(* IEC 61131-3 sources: daoli-st-library/DL_Process (part 67) *)

(* ---- FB_DL_ModbusPollMaster.st ---- *)
(*==============================================================================
 * 组件名称 (Component)  : FB_DL_ModbusPollMaster
 * 所属子库 (Sublibrary) : DL_Process
 * 当前版本 (Version)    : 1.0.0
 * 分类     (Category)   : 通信调度功能块（Function Block · 轮询主站调度抽象层）
 * 作者     (Author)     : Daoli Library
 * 日期     (Date)       : 2026-11-15
 * 兼容性   (Platform)   : CODESYS 3.5 / TwinCAT 3 / 汇川 InoProShop / Schneider
 *                         Machine Expert；纯 IEC 61131-3（第 3 版）语法，
 *                         仅依赖 Standard.library（TON / F_TRIG），零厂商方言
 * 功能简介 (Function)   : 多从站轮询主站调度器（Modbus RTU 轮询节拍抽象层）。
 *                         按站表顺序轮询、单事务响应超时重试、成功/异常双计数器
 *                         台账、空表与全跳过保护、站表禁用跳过的自动回绕。本块
 *                         只做「调度」：决定「此刻该问哪个站、问什么地址区、失败
 *                         重试几次、超时怎么记账」，帧的构造、CRC 校验、字节收发、
 *                         串口/TCP 底层时序全部交由传输层实现。
 * 分层声明 (Layering)   : ① 本块不绑定任何具体串口库、不引用任何厂商驱动块；
 *                         ② 传输层经两个抽象方法 SendFrame / RecvFrame 由集成者
 *                         实现（推荐做法：EXTENDS 本块并覆盖 DoTransaction 作为
 *                         统一入口，在覆盖体内调用自家收发库，再复用本块的记账
 *                         与重试；亦可只覆盖 SendFrame / RecvFrame 两个帧级原语）；
 *                         ③ 基类默认实现为「抽象桩」：返回 FALSE 并锁故障码
 *                         0005_0290（传输层未实现），这是抽象层的合法形态，不是
 *                         漏填——未注入传输层时块不会静默假成功；
 *                         ④ 调度层零触碰帧内容：不解析功能码、不读写应答字节、
 *                         不做 CRC 运算。CRC-16/Modbus 的公开算法定义在本库已有
 *                         实现（见 DL_MathData 子库既有 CRC 计算函数），本块仅在
 *                         此注释说明「可作校验实现」，不 import、不调用、不内联。
 * 职责边界 (Scope)      : ① 不做站内数据解包与工程量换算（由上层按站表项自行
 *                         读取应答缓冲后处理）；② 不做主备链路切换与总线诊断
 *                         （后续轮次另立组件）；③ 不做写单寄存器/写多寄存器的
 *                         流程编排（功能码仅作透传字段，调度节拍与读写无关）。
 * 开源溯源 (Origin)     : 来源标签 codesys-forge-modbus（T1-4 开族续挖）。仅参考
 *                         CODESYS Forge 免费库 ModbusFB 公开文档页中「主站轮询 /
 *                         站表组织 / 超时重试 / 轮询间隔」的功能分类与参数域惯例，
 *                         以及「帧构造与校验归传输层」的分层语义；所据页面未显
 *                         式声明许可条款，故按最严口径处置：只借组织分类与参数
 *                         范围，零代码行复制。本块的枚举编号、状态机、站表结构、
 *                         台账口径与故障码位 100% 本库独立设计，clean-room 实现。
 * 公约遵循 (Convention) : 0.1/R19 首扫范式（IF (NOT _bInit)）；0.2/R21 bError 显式
 *                         排除信息级码；0.5/R7 定时器与边沿实例主体最前部无条件
 *                         刷新；0.6/R14 定时器语义参数变化断输入一拍；0.7/R15 故障
 *                         级锁存仅重建路径清码；0.9 出口默认值先赋；0.14 WHILE 带
 *                         防死锁计数器 + 数组访问先判上下界；0.16 阈值全常量化。
 * 红线自检 (Redline)    : 全局隔离 ✓（零全局变量表引用、零外部变量声明、零物理
 *                         地址字面记号）｜命名合规 ✓（b/n/u/f/t/a/st/e/fb/i 前缀
 *                         全覆盖）｜注释完整 ✓（声明行 100% 中英双语同行注释）｜
 *                         OOP 封装 ✓（内部状态全私有，传输层经抽象方法注入）｜
 *                         周期安全 ✓（TON / F_TRIG 实例无条件刷新，方法无跨周期
 *                         驻留）｜防御编程 ✓（索引判界、循环防死锁、重试上限、
 *                         ENUM + CASE + ELSE 兜底）｜可移植性 ✓（纯 IEC 61131-3）｜
 *                         终结符成对 ✓
 * 设计要点 (Key notes)  : ① 事务生命周期：eRequest 发起（一次性调用抽象方法）→
 *                         eWaitResp 轮询结果（ePending 等待、eDone 成功、
 *                         eTimeout/eFailed 失败）→ eSttUpdate 记账 → eNextStn。
 *                         传输层可为异步（返回 FALSE 且 eResult = ePending 表示
 *                         尚未收完），调度层的响应超时定时器是它的兜底下限。
 *                         ② 不因单站失败中断轮询：重试耗尽只累加该站异常计数并
 *                         继续下一站（台账留证，避免一站坏总线导致全线停摆）；
 *                         只有「传输层未实现」与「站表索引越界」才锁全局故障。
 *                         ③ 轮询间隔由 TON 闸门实现（eSttUpdate 后重新计时），
 *                         事务结束到下一次发起至少间隔 tPollInterval，防止从站
 *                         换向静默期被打断（RTU 帧间静默的工程近似）。
 *                         ④ 站表回绕：每次事务结束把索引 +1，寻找下一站时从当前
 *                         索引起最多检查 uStationCount 站（超过即回绕），全部
 *                         跳过则置信息级码并按间隔节流空转，不锁故障。
 *                         ⑤ 计数口径：uStatOk / uStatErr 累计在调用方持有的站表
 *                         项内（跨班不清零），本块自身不保存历史，重启即从站表
 *                         现值继续，便于 HMI 做长期台账。
 * 偏离留档 (Deviation)  : ① 规格建议故障码 0005_0290~0293 中 0293 未使用（站数
 *                         非法按钳位 + 信息级处置，不锁故障；理由：站数是可在线
 *                         修改的组态量，钳位比停机更符合现场），实际使用
 *                         0005_0290~0292 三条；
 *                         ② 传输层抽象未采用独立 INTERFACE 文件（理由：本库公约
 *                         0.18「一文件一 POU」，接口件须独立成 .st 且本泳道不
 *                         允许新增第 6 个文件；改为块内抽象方法三件套，语义等价：
 *                         基类桩返回 FALSE + 锁码，派生块覆盖实现）；
 *                         ③ 规格 VAR 段 bFirstScan 改名 _bInit（公约 0.1 统一命名）。
 * 故障码表 (Error codes) :
 *                         16#0005_0190【信息级】站数越界已钳位到 1 至 16
 *                         16#0005_0191【信息级】站表全部跳过，本轮无事务（按间隔节流）
 *                         16#0005_0192【信息级】单站重试耗尽，异常台账已累加
 *                         16#0005_0193【信息级】超时/间隔参数非法已兜底
 *                         16#0005_0290【故障级】传输层未实现（抽象方法桩未被覆盖）
 *                         16#0005_0291【故障级】站表索引越界（越界保护触发）
 *                         16#0005_0292【故障级】非法状态兜底（枚举越界）
 * 验收向量 (Acceptance) :
 *   V1 单站成功：站数 1、从站 1 功能码 3 → eRequest 发起一次，eWaitResp 得
 *      eDone → uStatOk +1、bDone 单拍、回到 eNextStn；
 *   V2 超时重试：传输层持续回 ePending → 响应超时定时器到期后 uActiveRetry
 *      逐次 +1，达 uMaxRetry 后该站 uStatErr +1 且轮询继续下一站（不锁故障）；
 *   V3 站表跳过：站 0 的 bSkip = TRUE → 首个事务直接落在站 1（索引回绕正确）；
 *      全部站跳过 → 信息级 0191，块按 tPollInterval 节流空转，bBusy FALSE；
 *   V4 抽象桩：未覆盖 DoTransaction / SendFrame / RecvFrame → 首次发起即锁
 *      0005_0290 并停轮询，bError TRUE（杜绝静默假成功）；
 *   V5 间隔节流：tPollInterval = 100 ms、任务 10 ms → 相邻两事务发起间隔
 *      不少于 100 ms（TON 闸门计时）；
 *   V6 禁用重建：bEnable 下降沿 → 队伍暂停且保持现场（站索引/计数不清零），
 *      再次使能从原索引继续，不重复打扰刚问过的站。
 * 修订历史 (Revision)   :
 *   2026-11-15  v1.0.0  首版入库（Round 09 · DL_Process Modbus 轮询调度件）
 *============================================================================*)

(*-----------------------------------------------------------------------------
 * 集成示例 (Integration guide)：
 *   1 定义派生块 FB_MyRtuMaster EXTENDS FB_DL_ModbusPollMaster，覆盖
 *     DoTransaction（VAR_IN_OUT stItem : ST_DL_PollItem），在覆盖体内调用自家
 *     串口收发块完成「组帧 + 发送 + 收帧 + CRC 校验」，并把结果写回本块事务
 *     上下文（成功回 eDone，超时回 eTimeout，异常码回 uExceptionCode）。
 *   2 上层每周期调用派生块实例，注入站表数组与调度参数：
 *      aPollTable[0].uSlaveAddr := 1; aPollTable[0].uFuncCode := 3;
 *      aPollTable[0].uStartAddr := 0; aPollTable[0].uQuantity := 16;
 *      fbPoll(uStationCount := 4, tRespTimeout := T#500MS, uMaxRetry := 3,
 *             tPollInterval := T#100MS, aPollTable := aPollTable);
 *   3 读台账：aPollTable[i].uStatOk / uStatErr 由本块维护，HMI 直接读结构体。
 *----------------------------------------------------------------------------*)

(*-----------------------------------------------------------------------------
 * 常见误用与现场提示 (Field notes)：
 *   1 站表项的功能码只是透传字段，本块不校验其合法性；上位填 0 或非法功能码
 *     时，从站会回异常码，表现为该站 uStatErr 持续上升，请查站表而不是本块。
 *   2 响应超时必须大于最慢从站的最长应答时间；填得过小会造成「其实成功但被
 *     判超时」的重复点名，从站可能因此回异常码（上一次未收完）。
 *   3 uMaxRetry = 0 表示不重试，一次失败即记账进下一站，适合「宁漏不拖」的
 *     快速巡检场景。
 *   4 站表全部 bSkip 时本块按间隔空转且 bBusy 恒 FALSE，这是正常状态，不是
 *     死机；检修期整线隔离时常被误判为故障。
 *   5 本块不做总线抢占仲裁：同一物理链路上不要挂两个本块实例，否则帧会交错。
 *----------------------------------------------------------------------------*)

(*-----------------------------------------------------------------------------
 * 枚举: E_DL_PollState（归属 FB_DL_ModbusPollMaster，随本文件发布）
 * 含义: 轮询调度离散状态。数值步长 10 留空位，故障态 99 保证排序末位。
 *----------------------------------------------------------------------------*)
{attribute 'strict'}
{attribute 'qualified_only'}
TYPE E_DL_PollState :
(
    eIdle      := 0,     // 空闲：未使能或故障重建后待启动 / Idle: disabled or waiting for a rebuild
    eNextStn   := 10,    // 选下一站：按站表回绕寻找未跳过站，并受轮询间隔闸门约束 / Select next station with wrap and interval gating
    eRequest   := 20,    // 发起事务：一次性调用抽象方法 DoTransaction / Issue one transaction by calling DoTransaction
    eWaitResp  := 30,    // 等待应答：轮询传输层结果与响应超时定时器 / Wait for the transport result and the response timeout
    eSttUpdate := 40,    // 记账：成功/异常计数累加并产生单拍完成脉冲 / Accounting with a one-scan done pulse
    eFault     := 99     // 故障锁存：仅使能下降沿重建可退 / Fault latched, left only by the disable-edge rebuild
) UINT;
END_TYPE

(*-----------------------------------------------------------------------------
 * 枚举: E_DL_MbTxnResult（归属 FB_DL_ModbusPollMaster，随本文件发布）
 * 含义: 单事务结果，由传输层回填。调度层只据此推进状态，不解析帧内容。
 *----------------------------------------------------------------------------*)
{attribute 'strict'}
{attribute 'qualified_only'}
TYPE E_DL_MbTxnResult :
(
    ePending := 0,       // 传输中：尚未收完应答（异步传输层的等待态） / In progress, response not yet complete
    eDone    := 10,      // 事务成功：应答完整且通过传输层校验 / Success, a complete and validated response
    eTimeout := 20,      // 传输超时：传输层自身判超时 / Timeout reported by the transport layer
    eFailed  := 30       // 传输失败：校验错、异常码或链路错误 / Failure such as a check error, an exception or a link error
) UINT;
END_TYPE

(*-----------------------------------------------------------------------------
 * 结构体: ST_DL_PollItem（归属 FB_DL_ModbusPollMaster，随本文件发布）
 * 用途: 站表项。由调用方持有并注入（VAR_IN_OUT 数组），本块只读写统计字段。
 * 说明: uFuncCode / uStartAddr / uQuantity 均为透传字段，本块不解析、不改写。
 *----------------------------------------------------------------------------*)
TYPE ST_DL_PollItem :
STRUCT
    uSlaveAddr : USINT := 1;      // 从站地址（Slave address）[1~247]，0 与 248 以上为保留地址 / Reserved above 247 and at zero
    uFuncCode  : USINT := 3;      // 功能码（Function code），本块仅透传不解析 / Passed through, never parsed by this block
    uStartAddr : UINT := 0;       // 起始地址（Start address），寄存器区偏移，本块仅透传 / Register offset, passed through only
    uQuantity  : UINT := 1;       // 数量（Quantity），寄存器个数或线圈个数，本块仅透传 / Register or coil count, passed through only
    uStatOk    : UDINT := 0;      // 成功计数（Success counter）[次]，跨班累计由调用方清零 / Accumulated until the caller clears it
    uStatErr   : UDINT := 0;      // 异常计数（Error counter）[次]，重试耗尽即累加 / Incremented when the retries are exhausted
    bSkip      : BOOL := FALSE;   // 本站跳过（Skip this station），TRUE 时轮询回绕绕过本站 / TRUE makes the scan wrap past this station
END_STRUCT
END_TYPE

(*-----------------------------------------------------------------------------
 * 结构体: ST_DL_ModbusTxn（归属 FB_DL_ModbusPollMaster，随本文件发布）
 * 用途: 单事务上下文。调度层装填请求字段，传输层回填结果字段，双方以此交接。
 * 说明: 应答缓冲容量 256 字节为 Modbus RTU 最大帧长度（地址 + 功能码 + 数据 +
 *       CRC 的上限），调度层只保存不解读。
 *----------------------------------------------------------------------------*)
TYPE ST_DL_ModbusTxn :
STRUCT
    uSlaveAddr     : USINT := 1;                        // 从站地址（Slave address）[1~247] / Slave address in the range one to 247
    uFuncCode      : USINT := 3;                        // 功能码（Function code），透传 / Passed-through function code
    uStartAddr     : UINT := 0;                         // 起始地址（Start address），透传 / Passed-through start address
    uQuantity      : UINT := 1;                         // 数量（Quantity），透传 / Passed-through quantity
    eResult        : E_DL_MbTxnResult := E_DL_MbTxnResult.ePending; // 事务结果（Transaction result），传输层回填 / Filled in by the transport layer
    uExceptionCode : USINT := 0;                        // 异常码（Exception code）[1~255]，0 = 无异常，传输层回填 / Zero means no exception
    uRxLen         : UINT := 0;                         // 应答字节数（Response length）[字节]，传输层回填 / Response length in bytes
    auRxFrame      : ARRAY[0..255] OF BYTE;             // 应答帧原始字节（Raw response frame）[字节]，容量 256，调度层不解读 / Raw bytes, never parsed here
    bAbort         : BOOL := FALSE;                     // 中止请求（Abort request），重试或切站时由调度层置位 / Set by the scheduler on retries
END_STRUCT
END_TYPE

(*==============================================================================
 * 功能块: FB_DL_ModbusPollMaster
 * 调用约定: 每个扫描周期无条件调用一次；站表与参数全部经引脚注入。
 * 抽象层形态: DoTransaction / SendFrame / RecvFrame 三个默认实现均为抽象桩
 *             （返回 FALSE 并锁 0005_0290），由派生块覆盖后落地真实传输。
 *============================================================================*)
FUNCTION_BLOCK FB_DL_ModbusPollMaster
VAR_INPUT
    bEnable       : BOOL;               // 调度使能（Scheduler enable），FALSE 时队列暂停并保持现场 / FALSE pauses the queue and keeps the context
    uStationCount : UINT := 4;          // 轮询站数（Station count）[站]，域 1~16，越界钳位 / Clamped to the range one to sixteen
    tRespTimeout  : TIME := T#500MS;    // 单事务响应超时（Response timeout）[ms]，域 >= 1 ms / At least one millisecond
    uMaxRetry     : UINT := 3;          // 超时重试上限（Retry limit）[次]，0 = 不重试 / Zero means no retry
    tPollInterval : TIME := T#100MS;    // 相邻事务最小间隔（Minimum poll interval）[ms]，0 = 不节流 / Zero disables the interval gate
END_VAR
VAR_OUTPUT
    bBusy          : BOOL;              // 有事务执行中（Transaction in progress）/ A transaction is running
    uActiveStation : UINT;              // 当前轮询站索引（Active station index）[索引 0~15] / Active station index in the range zero to fifteen
    uActiveRetry   : UINT;              // 当前站累计重试数（Active retry count）[次]，切站清零 / Cleared when the station advances
    bDone          : BOOL;              // 单站事务完成（Station transaction done），单拍脉冲（R25）/ One-scan pulse per station completion
    bError         : BOOL;              // 故障保持型（Fault latched），显式排除信息级码 / Latched fault flag, info codes excluded
    uErrorId       : UDINT;             // 故障码（Error code），0 = 无故障，段位 16#0005_xxxx / Error code, zero means no error
END_VAR
VAR_IN_OUT
    aPollTable    : ARRAY[0..DL_MB_MAX_STN-1] OF ST_DL_PollItem; // 轮询站表（Poll table），调用方持有 / Caller-owned poll table
END_VAR
VAR
    _eState       : E_DL_PollState := E_DL_PollState.eIdle; // 主状态机状态（Main state machine state）/ Main state machine state
    _bInit        : BOOL;               // 首扫完成标志（First-scan done flag），初值 FALSE / First-scan done flag, initial FALSE
    _uStnIdx      : UINT;               // 当前站索引（Current station index）[索引]，域 0~15 / Station index in the range zero to fifteen
    _uRetryCnt    : UINT;               // 重试计数（Retry counter）[次] / Retry counter
    _uStnCntEff   : UINT := 4;          // 生效站数（Effective station count）[站]，钳位后 / Effective station count after clamping
    _uStnTried    : UINT;               // 已检查站数（Stations examined）[站]，回绕寻找用 / Stations examined during the wrap search
    _uGuard       : UINT;               // 循环防死锁计数（Loop guard counter）[次]，上限 16 / Loop guard bounded by sixteen
    _bStationFound : BOOL;              // 找到可轮询站（Usable station found）/ A usable station was found
    _tRespEff     : TIME := T#500MS;    // 生效响应超时（Effective response timeout）[ms] / Effective response timeout [ms]
    _tGapEff      : TIME := T#100MS;    // 生效轮询间隔（Effective poll interval）[ms] / Effective poll interval [ms]
    _bGapActive   : BOOL;               // 间隔闸门激活（Interval gate armed），TRUE 时须等定时器到期 / The gate holds until the timer elapses
    _bGapBreak    : BOOL;               // 间隔定时器断输入一拍（Interval timer break），重新计时用（公约 0.6）/ One-scan break used to restart the timer
    _bGapFeed     : BOOL;               // 间隔定时器输入（Interval timer input），先算后喂（公约 0.5）/ Computed first and then fed to the timer
    _bRespBreak   : BOOL;               // 超时定时器断输入一拍（Timeout timer break），发起事务后重计时 / One-scan break after a request is issued
    _bRespFeed    : BOOL;               // 超时定时器输入（Timeout timer input），先算后喂（公约 0.5）/ Computed first and then fed to the timer
    _stTxn        : ST_DL_ModbusTxn;    // 事务上下文（Transaction context），与传输层交接 / Transaction context shared with the transport
    _bTxnOk       : BOOL;               // 本次事务成功（Transaction succeeded）/ Transaction succeeded flag
    _bTxnStub     : BOOL;               // 抽象方法桩未覆盖（Stub not overridden），TRUE 即锁故障 / TRUE when the abstract stub is still in place
    _bFaultLatch  : BOOL;               // 故障锁存（Fault latch），仅重建路径清除 / Fault latch, cleared only through the rebuild path
    _uErrInt      : UDINT;              // 故障级码寄存（Fault-level code register），锁存型 / Latched fault-level code register
    _uInfoCode    : UDINT;              // 本拍信息级码（Info code this scan），每拍重算 / Info code recomputed every scan
    _fbPollTick   : TON;                // 轮询间隔定时器（Poll interval timer），主周期无条件刷新 / Refreshed unconditionally every scan
    _fbRespWatch  : TON;                // 响应超时定时器（Response watchdog timer），主周期无条件刷新 / Refreshed unconditionally every scan
    _fbTrigDisable : F_TRIG;            // 使能下降沿（Enable falling edge），故障重建触发 / Triggers the disable-edge rebuild
END_VAR
VAR CONSTANT
    DL_MB_MAX_STN  : UINT := 16;        // 最大站数（Maximum station count）[站]，同时为站表长度 / Maximum station count, also the table length
    DL_MB_FRAME_MAX : UINT := 256;      // 最大帧长（Maximum frame length）[字节]，Modbus RTU 上限 / Modbus RTU frame limit
    DL_MAX_LOOP    : UINT := 16;        // 循环防死锁上限（Loop guard bound）[次]，等于站数上限 / Loop guard bound equal to the station limit
    DL_TIME_MIN    : TIME := T#1MS;     // 时间参数下限（Lower time bound）[ms]，兜底用 / Lower bound used when a time input is illegal
    DL_STN_MIN     : UINT := 1;         // 站数下限（Lower station bound）[站] / Lower bound of the station count
END_VAR

METHOD DoTransaction : BOOL
VAR_IN_OUT
    stItem : ST_DL_PollItem;           // 站表项（Poll item），只读意图，统计字段由主体维护 / Read-only intent, statistics maintained by the body
END_VAR
_stTxn.uSlaveAddr     := stItem.uSlaveAddr; // 装填从站地址（Fill the slave address）
_stTxn.uFuncCode      := stItem.uFuncCode;  // 装填功能码（Fill the function code）
_stTxn.uStartAddr     := stItem.uStartAddr; // 装填起始地址（Fill the start address）
_stTxn.uQuantity      := stItem.uQuantity;  // 装填数量（Fill the quantity）
_stTxn.eResult        := E_DL_MbTxnResult.ePending; // 结果置等待态（Result set to pending）
_stTxn.uExceptionCode := 0;                 // 异常码清零（Exception code cleared）
_stTxn.uRxLen         := 0;                 // 应答长度清零（Response length cleared）
IF SendFrame(stTxn := _stTxn) THEN
    IF RecvFrame(stTxn := _stTxn) THEN
        _stTxn.eResult := E_DL_MbTxnResult.eDone; // 收帧完成即置成功（A complete response marks success）
    END_IF
ELSIF NOT _bTxnStub THEN
    _stTxn.eResult := E_DL_MbTxnResult.eFailed; // 发送失败且非桩未覆盖（Send failure, not the stub case）
END_IF
DoTransaction := (_stTxn.eResult = E_DL_MbTxnResult.eDone); // 仅成功返回 TRUE（TRUE only on success）

(*------------------------------------------------------------------------------
 * 方法: SendFrame —— 帧级发送原语（抽象桩）。派生块覆盖后在体内完成组帧与发送。
 *      Method SendFrame - frame level transmit primitive, an abstract stub here.
 *------------------------------------------------------------------------------*)
    END_METHOD

METHOD SendFrame : BOOL
VAR_IN_OUT
    stTxn : ST_DL_ModbusTxn;           // 事务上下文（Transaction context），承载请求字段与中止标志 / Carries the request fields and the abort flag
END_VAR
IF stTxn.bAbort THEN
    stTxn.eResult := E_DL_MbTxnResult.eFailed; // 已请求中止则不再发送（Aborted transactions are not transmitted）
    SendFrame     := FALSE;            // 未发送（Not transmitted）
ELSE
    _bTxnStub := TRUE;                 // 标记抽象桩未被覆盖（Mark the stub as not overridden）
    SendFrame := FALSE;                // 桩一律返回 FALSE（The stub always returns FALSE）
END_IF

(*------------------------------------------------------------------------------
 * 方法: RecvFrame —— 帧级接收原语（抽象桩）。派生块覆盖后在体内完成收帧与校验。
 *      Method RecvFrame - frame level receive primitive, an abstract stub here.
 *------------------------------------------------------------------------------*)
    END_METHOD

METHOD RecvFrame : BOOL
VAR_IN_OUT
    stTxn : ST_DL_ModbusTxn;           // 事务上下文（Transaction context），承载结果字段回填 / Carries the result fields to be filled in
END_VAR
IF stTxn.bAbort THEN
    stTxn.eResult := E_DL_MbTxnResult.eFailed; // 已请求中止则不收帧（Aborted transactions are not received）
    RecvFrame     := FALSE;            // 未接收（Not received）
ELSE
    _bTxnStub := TRUE;                 // 标记抽象桩未被覆盖（Mark the stub as not overridden）
    RecvFrame := FALSE;                // 桩一律返回 FALSE（The stub always returns FALSE）
END_IF
    END_METHOD

// ============================================================================
// 段 1｜输出确定性默认值先赋（公约 0.9；R25 第一律：单拍标志每拍预清零）
//      Deterministic defaults first, one-scan flags pre-cleared every scan
// ============================================================================
bDone      := FALSE;                   // 完成脉冲预清零，仅 eSttUpdate 拍置位（Done pulse pre-cleared, set only in the update state）
bBusy      := FALSE;                   // 忙碌标志预清零（Busy flag pre-cleared）
_uInfoCode := 0;                       // 信息级码每拍重算（Info code recomputed every scan）

// ============================================================================
// 段 2｜首扫初始化（R19 范式）
//      First-scan initialization following the single legal R19 predicate
// ============================================================================
IF NOT _bInit THEN
    _bInit        := TRUE;             // 置首扫完成（First-scan done）
    _eState       := E_DL_PollState.eIdle; // 状态复位为空闲（State reset to idle）
    _uStnIdx      := 0;                // 站索引清零（Station index cleared）
    _uRetryCnt    := 0;                // 重试计数清零（Retry counter cleared）
    _bGapActive   := FALSE;            // 间隔闸门关闭（Interval gate disarmed）
    _stTxn.bAbort := FALSE;            // 事务中止标志清零（Transaction abort cleared）
    _bFaultLatch  := FALSE;            // 故障锁存清零（Fault latch cleared）
    _uErrInt      := 16#0000_0000;     // 故障码清零（Fault code cleared）
END_IF

// ============================================================================
// 段 3｜定时器与边沿实例无条件周期刷新（公约 0.5 / 0.6：入参先算后喂）
//      Unconditional refresh of timers and the edge instance
// ============================================================================
_fbTrigDisable(CLK := bEnable);        // 使能下降沿检测（Enable falling edge detection）

_bGapFeed := _bGapActive AND (NOT _bGapBreak); // 间隔定时器输入（Interval timer input）
_fbPollTick(IN := _bGapFeed, PT := _tGapEff);  // 间隔计时（Interval timing）
_bGapBreak := FALSE;                   // 断输入脉冲在实例调用后自清（Break pulse self-cleared after the call）

IF _fbPollTick.Q THEN
    _bGapActive := FALSE;              // 间隔已满，解除闸门（Gate released once the interval elapsed）
END_IF

_bRespFeed := (_eState = E_DL_PollState.eWaitResp) AND (NOT _bRespBreak); // 超时定时器输入（Timeout timer input）
_fbRespWatch(IN := _bRespFeed, PT := _tRespEff); // 响应超时计时（Response timeout timing）
_bRespBreak := FALSE;                  // 断输入脉冲自清（Break pulse self-cleared）

// ============================================================================
// 段 4｜参数钳位（站数 1~16、超时与间隔 >= 1 ms；越界只钳位并置信息级）
//      Parameter clamping, out-of-range values are clamped with info codes
// ============================================================================
IF uStationCount < DL_STN_MIN THEN
    _uStnCntEff := DL_STN_MIN;         // 站数下限钳位（Clamped to the lower bound）
    _uInfoCode  := 16#0005_0190;       // 0005_0190 站数越界已钳位【信息级】（Station count clamped, info level）
ELSIF uStationCount > DL_MB_MAX_STN THEN
    _uStnCntEff := DL_MB_MAX_STN;      // 站数上限钳位（Clamped to the upper bound）
    _uInfoCode  := 16#0005_0190;       // 0005_0190 站数越界已钳位【信息级】（Station count clamped, info level）
ELSE
    _uStnCntEff := uStationCount;      // 合法站数直通（Valid station count passed through）
END_IF

IF tRespTimeout < DL_TIME_MIN THEN
    _tRespEff  := DL_TIME_MIN;         // 超时下限兜底（Timeout falls back to the lower bound）
    _uInfoCode := 16#0005_0193;        // 0005_0193 超时/间隔参数非法已兜底【信息级】（Time parameter clamped, info level）
ELSE
    _tRespEff := tRespTimeout;         // 合法超时直通（Valid timeout passed through）
END_IF

IF tPollInterval = T#0MS THEN
    _tGapEff   := T#0MS;               // 间隔 0 = 不节流，定时器立即到期（Zero interval disables the gate, the timer expires at once）
    _uInfoCode := 16#0005_0193;        // 0005_0193 间隔参数为 0 已按不节流处置【信息级】（Zero interval treated as no gating, info level）
ELSE
    _tGapEff := tPollInterval;         // 合法间隔直通（Valid interval passed through）
END_IF

// ============================================================================
// 段 5｜站索引越界保护（防御性：正常流程不可达，纯兜底）
//      Station index guard, unreachable in the normal flow
// ============================================================================
IF _uStnIdx > DL_MB_MAX_STN THEN
    _bFaultLatch := TRUE;              // 索引越界锁故障（Out-of-range index latches a fault）
    _uErrInt     := 16#0005_0291;      // 0005_0291 站表索引越界【故障级】（Station index out of range, fault level）
    _uStnIdx     := 0;                 // 索引强制回零自愈（Index forced back to zero）
ELSIF _uStnIdx = DL_MB_MAX_STN THEN
    _uStnIdx := 0;                     // 恰在上界即回绕，属正常（Wrapping at the bound is the normal path）
END_IF

// ============================================================================
// 段 6｜主状态机（ENUM + CASE + ELSE 兜底；故障重建走使能下降沿）
//      Main state machine with mandatory ELSE fallback and a disable-edge rebuild
// ============================================================================
CASE _eState OF

    E_DL_PollState.eIdle: // 空闲：等使能（Idle, waiting for enable）
        IF _fbTrigDisable.Q THEN
            _bFaultLatch := FALSE;     // 下降沿重建：清故障锁存（Rebuild clears the fault latch）
            _uErrInt     := 16#0000_0000; // 故障码清零（Fault code cleared）
            _uRetryCnt   := 0;         // 重试计数清零（Retry counter cleared）
        END_IF
        IF bEnable AND (NOT _bFaultLatch) THEN
            _bGapActive := FALSE;      // 起动首事务不节流（The first transaction is not gated）
            _uRetryCnt  := 0;          // 重试计数清零（Retry counter cleared）
            _eState     := E_DL_PollState.eNextStn; // 进选站态（Enter the station selection state）
        END_IF

    E_DL_PollState.eNextStn: // 选下一站：回绕寻找 + 间隔闸门（Select next station with wrap and gating）
        IF (NOT bEnable) OR _bFaultLatch THEN
            _eState := E_DL_PollState.eIdle; // 使能撤销或故障即回空闲（Disabled or faulty returns to idle）
        ELSIF (NOT _bGapActive) OR _fbPollTick.Q THEN
            _bStationFound := FALSE;   // 站发现标志预清零（Station found flag pre-cleared）
            _uStnTried     := 0;       // 已检查站数清零（Stations examined cleared）
            _uGuard        := 0;       // 循环守卫清零（Loop guard cleared）
            WHILE (_uStnTried < _uStnCntEff) AND (_uGuard < DL_MAX_LOOP) AND (NOT _bStationFound) DO
                _uGuard    := _uGuard + 1;      // 循环守卫递增，防死锁（Guard incremented to prevent a dead loop）
                _uStnTried := _uStnTried + 1;   // 已检查站数递增（Stations examined incremented）
                IF _uStnIdx >= _uStnCntEff THEN
                    _uStnIdx := 0;              // 回绕到首站（Wrap back to the first station）
                END_IF
                IF NOT aPollTable[_uStnIdx].bSkip THEN
                    _bStationFound := TRUE;     // 找到可用站（Usable station found）
                ELSE
                    _uStnIdx := _uStnIdx + 1;   // 跳过本站，索引后移（Skip this station and advance）
                END_IF
            END_WHILE
            IF _bStationFound THEN
                _uRetryCnt  := 0;              // 新站重试计数清零（Retry counter cleared for the new station）
                _bRespBreak := TRUE;           // 超时定时器下拍从零开始（Timeout timer restarts next scan）
                _eState     := E_DL_PollState.eRequest; // 进发起态（Enter the request state）
            ELSE
                _uInfoCode  := 16#0005_0191;   // 0005_0191 站表全部跳过【信息级】（All stations skipped, info level）
                _bGapActive := TRUE;           // 按间隔节流空转（Idle pacing through the interval gate）
                _bGapBreak  := TRUE;           // 间隔定时器重新计时（Interval timer restarted）
            END_IF
        END_IF

    E_DL_PollState.eRequest: // 发起事务：一次性调用抽象方法（Issue one transaction）
        _stTxn.uSlaveAddr     := aPollTable[_uStnIdx].uSlaveAddr; // 透传从站地址（Pass the slave address through）
        _stTxn.uFuncCode      := aPollTable[_uStnIdx].uFuncCode;  // 透传功能码（Pass the function code through）
        _stTxn.uStartAddr     := aPollTable[_uStnIdx].uStartAddr; // 透传起始地址（Pass the start address through）
        _stTxn.uQuantity      := aPollTable[_uStnIdx].uQuantity;  // 透传数量（Pass the quantity through）
        _stTxn.eResult        := E_DL_MbTxnResult.ePending;       // 结果置等待态（Result set to pending）
        _stTxn.uExceptionCode := 0;                               // 异常码清零（Exception code cleared）
        _stTxn.uRxLen         := 0;                               // 应答长度清零（Response length cleared）
        _stTxn.bAbort         := FALSE;                           // 中止标志清零（Abort cleared）
        _bTxnStub             := FALSE;                           // 桩标志预清零（Stub flag pre-cleared）
        _bTxnOk               := DoTransaction(stItem := aPollTable[_uStnIdx]); // 抽象方法调用，每拍至多一次（At most one call per scan）
        _bRespBreak           := TRUE;                            // 超时定时器下拍从零开始（Timeout timer restarts next scan）
        IF _bTxnStub THEN
            _bFaultLatch := TRUE;        // 传输层未实现即锁故障（A missing transport latches a fault）
            _uErrInt     := 16#0005_0290; // 0005_0290 传输层未实现【故障级】（Transport not implemented, fault level）
            _eState      := E_DL_PollState.eFault;
        ELSE
            _eState := E_DL_PollState.eWaitResp; // 进等待应答态（Enter the waiting state）
        END_IF

    E_DL_PollState.eWaitResp: // 等待应答：结果枚举与超时定时器双判（Wait on the result and the watchdog）
        IF (_stTxn.eResult = E_DL_MbTxnResult.eDone) AND (_stTxn.uRxLen <= DL_MB_FRAME_MAX) THEN
            _bTxnOk := TRUE;             // 事务成功且帧长在容量内（Success with a length inside the buffer capacity）
            _eState := E_DL_PollState.eSttUpdate; // 进记账态（Enter the accounting state）
        ELSIF _stTxn.uRxLen > DL_MB_FRAME_MAX THEN
            _stTxn.bAbort := TRUE;       // 帧长越界即中止（Abort on an over-long frame）
            _bTxnOk := FALSE;            // 帧长越界判失败，不再重试（Over-long frame fails without a retry）
            _eState := E_DL_PollState.eSttUpdate; // 进记账态（Enter the accounting state）
        ELSIF (_stTxn.eResult = E_DL_MbTxnResult.eTimeout) OR
              (_stTxn.eResult = E_DL_MbTxnResult.eFailed) OR _fbRespWatch.Q THEN
            _stTxn.bAbort := TRUE;       // 通知传输层中止本事务（Ask the transport to abort）
            IF _uRetryCnt < uMaxRetry THEN
                _uRetryCnt := _uRetryCnt + 1;   // 重试计数累加（Retry counter incremented）
                _eState    := E_DL_PollState.eRequest; // 重新发起（Reissue the transaction）
            ELSE
                _bTxnOk := FALSE;        // 重试耗尽判失败（Retries exhausted, marked as failed）
                _eState := E_DL_PollState.eSttUpdate; // 进记账态（Enter the accounting state）
            END_IF
        END_IF

    E_DL_PollState.eSttUpdate: // 记账：台账累加 + 单拍完成脉冲 + 推进站索引（Accounting and advance）
        IF _bTxnOk THEN
            aPollTable[_uStnIdx].uStatOk := aPollTable[_uStnIdx].uStatOk + 1; // 成功计数累加（Success counter incremented）
        ELSE
            aPollTable[_uStnIdx].uStatErr := aPollTable[_uStnIdx].uStatErr + 1; // 异常计数累加（Error counter incremented）
            _uInfoCode := 16#0005_0192; // 0005_0192 单站重试耗尽【信息级】（Station retries exhausted, info level）
        END_IF
        bDone       := TRUE;           // 单站完成单拍脉冲，本拍不再清除（One-scan done pulse, never cleared in the same scan）
        _uRetryCnt  := 0;              // 切站重试计数清零（Retry counter cleared on the station change）
        IF (_uStnIdx + 1) >= _uStnCntEff THEN
            _uStnIdx := 0;             // 到表尾即回绕首站（Wrap to the first station at the table end）
        ELSE
            _uStnIdx := _uStnIdx + 1;  // 索引后移到下一站（Advance to the next station）
        END_IF
        _bGapActive := TRUE;           // 启用间隔闸门（Arm the interval gate）
        _bGapBreak  := TRUE;           // 间隔定时器重新计时（Interval timer restarted）
        _eState     := E_DL_PollState.eNextStn; // 回选站态（Back to the selection state）

    E_DL_PollState.eFault: // 故障锁存：停轮询，保持现场（Fault latched, polling stopped）
        IF _fbTrigDisable.Q THEN
            _bFaultLatch := FALSE;     // 使能下降沿重建（Rebuild on the enable falling edge）
            _uErrInt     := 16#0000_0000; // 故障码清零（Fault code cleared）
            _uRetryCnt   := 0;         // 重试计数清零（Retry counter cleared）
            _eState      := E_DL_PollState.eIdle; // 回空闲（Back to idle）
        END_IF

    ELSE
        _bFaultLatch := TRUE;          // 非法状态兜底锁存（Illegal state latched）
        _uErrInt     := 16#0005_0292;  // 0005_0292 非法状态兜底【故障级】（Illegal state fallback, fault level）
        _eState      := E_DL_PollState.eFault; // 进故障态（Enter the fault state）
END_CASE

// ============================================================================
// 段 7｜出口映射（忙碌派生、活动站索引、重试数、故障级码优先透出）
//      Outlet mapping with fault-level codes taking priority over info codes
// ============================================================================
bBusy          := (_eState = E_DL_PollState.eRequest) OR (_eState = E_DL_PollState.eWaitResp); // 忙碌派生（Busy derived form）
uActiveStation := _uStnIdx;            // 活动站索引出口（Active station index outlet）
uActiveRetry   := _uRetryCnt;          // 活动重试数出口（Active retry count outlet）
bError         := _bFaultLatch OR (_eState = E_DL_PollState.eFault); // 故障派生，显式排除信息级（Fault derived, info codes excluded）
IF bError THEN
    uErrorId := _uErrInt;              // 故障级码优先（Fault-level code has priority）
ELSE
    uErrorId := _uInfoCode;            // 无故障透出本拍信息级码（Transient info code exposed）
END_IF

(*------------------------------------------------------------------------------
 * 方法: DoTransaction —— 抽象入口：装填上下文、调用帧级原语、返回成功与否。
 *      Method DoTransaction - abstract entry assembling the context and calling
 *      the frame level primitives. Derived blocks override this method.
 *------------------------------------------------------------------------------*)

END_FUNCTION_BLOCK

(* ---- FB_DL_ModulePottingVac.st ---- *)
(*==============================================================================
 * 组件名称 (Component)  : FB_DL_ModulePottingVac
 * 所属子库 (Sublibrary) : DL_Process
 * 当前版本 (Version)    : 1.0.1
 * 兼容性   (Platform)   : CODESYS 3.5+ / TwinCAT 3 / 汇川 InoProShop / 施耐德 Machine Expert
 *                         仅依赖 Standard.library（TON / R_TRIG），零厂商私有库
 * 功能描述 (Function)   : 灌胶真空脱泡四相顺控：抽真空 → 保持 → 破空 → 泄压。
 *                         每相一个**专用** TON，PT 语义各自成对写死，绝不共用一个实例改 PT：
 *                           eEvac   抽真空：tonEvacTo  PT = tEvac    （到真空位 bVacReached 即过相）
 *                           eHold   保持  ：tonHoldTo  PT = tHold    （纯定时过相，无外部条件）
 *                           eBreak  破空  ：tonBreakTo PT = tBreak   （到常压位 bBreakDone 即过相）
 *                           eRelief 泄压  ：tonReliefTo PT = tRelief （纯定时过相，完成后回 eIdle）
 *                         每相的"过相条件"= 定时到 ∧ 该相到位信号（有到位信号的两相）；定时到但
 *                         到位信号没来 = 该相超时 → eFault（归因按相区分：eVacTimeout /
 *                         eBreakTimeout）。保持相与泄压相无到位信号，定时到即过相。
 *                         **eFault 可迁出**：bReset 上升沿 → 回 eIdle 并清 _eFaultFrom；同时 eFault
 *                         记录"从哪一相跌进故障"（_eFaultFrom），供 HMI 指明卡在哪一步。
 *                         bStop 在任一相立即可用 → 回 eIdle（中止，bAborted 单拍脉冲），中途中止
 *                         不记故障（操作员主动停机不是故障）。
 * 接口     (Interface)  : 输入 bStart 启动沿、bStop 中止、bVacReached 真空到位、bBreakDone 破空
 *                         到位、四相时间 tEvac / tHold / tBreak / tRelief、bReset 故障复位；
 *                         输出 bEvacActive / bHoldActive / bBreakActive / bReliefActive 四相指示、
 *                         bBusy 顺控进行中、bComplete 完成单拍、bAborted 中止单拍、ePhase 当前相、
 *                         eFaultFrom 跌入故障的相、eCause 成因、bError 故障标志。
 * 边界     (Boundary)   : ① **属主边界（写死）：本件只做四相时序编排，不驱动真空泵/破空阀/
 *                         泄压阀线圈**。阀/泵动作由 IO 映射层与执行件（`I_DL_Cylinder` 族或
 *                         阀门件）负责；本件出相指示位，由上层映射到实际输出。
 *                         ② 组态闸：任一相时间 <= T#0S → 故障锁存（零时长会让相瞬间过相，
 *                         工艺上等于跳过该相，是危险默认）。
 *                         ③ 四枚专用超时 TON（tonEvacTo / tonHoldTo / tonBreakTo / tonReliefTo）
 *                         在段 0 **无条件周期调用**，IN 由"当前相"表达式派生：进相即计时、出相即
 *                         复位，因此不存在跨相累积（R228A：专用超时 TON 命名豁免 + IN 表达式派生）；
 *                         PT 各绑一个专用时间引脚，绝不复用实例改 PT。
 *                         ④ eFault 迁出链：bReset 上升沿 → eIdle（清 _eFaultFrom 与 _eCause）；
 *                         bStop 亦可在故障相把相序拉回 eIdle（停机优先于故障保持），两条路径
 *                         都在段 3 显式写出（R228B 可迁出）。
 *                         ⑤ 零全局耦合（无 GVL / 无 VAR_EXTERNAL / 无物理地址）。
 *                         ⑥ **到位信号沿锁存语义（v1.0.1 修订）**：bVacReached / bBreakDone 允许
 *                         为短脉冲型（如压力开关瞬时动作）——两路各设 R_TRIG（段 0 无条件刷新）
 *                         + 锁存量 _bVacSeen / _bBreakSeen，进相首拍清锁存、捕获到位沿后置位；
 *                         过相判据读锁存量（tonEvacTo.Q AND _bVacSeen），脉冲先于超时 TON 到 Q
 *                         消失不再误报超时；持续到位信号行为不变（契约兼容）；迁出链（复位沿 /
 *                         bStop）同时清两锁存量，防跨循环残留。
 * 分工声明 (Scope)      : 与 `FB_DL_PressureDecayTest` 一类气密测试件分工——那件判"密封性"
 *                         （压降速率），本件只管"四相走完没走完、有没有卡相"；不共用判据。
 * 来源标签 (Source Tag) : ROADMAP B 类 / T2-8（灌胶真空脱泡四相顺控，自研 clean-room）
 * 解除式   (Release)    : bReset 上升沿 ∨ bStop（停机优先）→ 回 eIdle 并清故障记录。
 *                         自证可满足：两个外部信号均为操作员级动作，不受任何锁存量门控；
 *                         不存在"必须先到某相才能复位"的隐含前置。
 * 码表     (Codes)      : 本件不占用任何全局数字码位。出口为 ENUM 相别 + ENUM 成因 + BOOL 组；
 *                         数字码位待主控收口阶段统一派号。
 * 红线自检 (Redline)    : R1 ✓ 零 GVL/VAR_EXTERNAL ｜ R2 ✓ 零 %I/%Q/%M ｜ R3 ✓ 纯 IEC 61131-3
 *                         R4 ✓ 时间域几何闸 + 无浮点比较 ｜ R5 ✓ 声明逐行同行双语注释
 *                         R6 ✓ ENUM+CASE 含 ELSE ｜ R7 ✓ 四 TON/两沿段 0 无条件刷新
 * 修订历史 (Revision)   : 2026-11-19  v1.0.0  R46 首版（批次 4 · 序号 19）
 *                         2026-11-20  v1.0.1  R47 终审轻项返修：到位脉冲先于超时 TON 到 Q 消失
 *                         导致过相判据恒假误报超时；增到位沿 R_TRIG 锁存 _bVacSeen/_bBreakSeen，
 *                         过相判据改读锁存量，迁出链清锁存；引脚契约零变更，V1~V3 向量保持。
 *==============================================================================*)

TYPE E_DL_MpvPhase :
(
    eIdle   := 0,    // 待机相 / Idle
    eEvac   := 10,   // 抽真空相 / Evacuation
    eHold   := 20,   // 真空保持相 / Vacuum hold
    eBreak  := 30,   // 破空相 / Air break
    eRelief := 40,   // 泄压相 / Pressure relief
    eFault  := 90    // 故障相（等复位） / Fault, awaiting reset
);
END_TYPE

TYPE E_DL_MpvCause :
(
    eNone         := 0,   // 无异常 / No anomaly
    eCfgIllegal   := 1,   // 组态非法（相时间非正） / Illegal configuration
    eVacTimeout   := 2,   // 抽真空相超时（未到真空位） / Evacuation timed out before reaching vacuum
    eBreakTimeout := 3,   // 破空相超时（未到常压位） / Air break timed out before reaching atmosphere
    ePhaseBad     := 4    // 非法相位兜底 / Illegal phase fallback
);
END_TYPE

FUNCTION_BLOCK FB_DL_ModulePottingVac
VAR_INPUT
    bStart      : BOOL := FALSE;        // 启动沿，进入抽真空相 [-] / Start edge, enters evacuation
    bStop       : BOOL := FALSE;        // 中止（停机优先，任一相可用） [-] / Abort, honoured in every phase
    bVacReached : BOOL := FALSE;        // 真空到位信号（抽真空相过相条件） [-] / Vacuum reached, evacuation exit condition
    bBreakDone  : BOOL := FALSE;        // 破空到位信号（破空相过相条件） [-] / Atmosphere reached, air-break exit condition
    tEvac       : TIME := T#30S;        // 抽真空相超时，域 > T#0S [ms] / Evacuation timeout, > T#0S [ms]
    tHold       : TIME := T#10S;        // 真空保持时长，域 > T#0S [ms] / Vacuum hold duration, > T#0S [ms]
    tBreak      : TIME := T#10S;        // 破空相超时，域 > T#0S [ms] / Air-break timeout, > T#0S [ms]
    tRelief     : TIME := T#5S;         // 泄压时长，域 > T#0S [ms] / Pressure-relief duration, > T#0S [ms]
    bReset      : BOOL := FALSE;        // 故障复位，上升沿回待机相 [-] / Fault reset, rising edge returns to idle
END_VAR
VAR_OUTPUT
    bEvacActive   : BOOL;               // 抽真空相进行中 [-] / Evacuation phase active
    bHoldActive   : BOOL;               // 真空保持相进行中 [-] / Hold phase active
    bBreakActive  : BOOL;               // 破空相进行中 [-] / Air-break phase active
    bReliefActive : BOOL;               // 泄压相进行中 [-] / Relief phase active
    bBusy         : BOOL;               // 顺控进行中（非待机非故障） [-] / Sequence busy
    bComplete     : BOOL;               // 四相完成，单拍脉冲 [-] / Sequence complete, single-scan pulse
    bAborted      : BOOL;               // 中止，单拍脉冲 [-] / Aborted, single-scan pulse
    ePhase        : E_DL_MpvPhase;      // 当前相出口 [-] / Present phase outlet
    eFaultFrom    : E_DL_MpvPhase;      // 跌入故障时所处的相（诊断用） [-] / Phase that faulted
    eCause        : E_DL_MpvCause;      // 成因出口（R190 归因唯一） [-] / Cause outlet
    bError        : BOOL;               // 故障标志（组态非法或相超时） [-] / Error flag
END_VAR
VAR
    _eState    : E_DL_MpvPhase := E_DL_MpvPhase.eIdle;    // 内部相（CASE 唯一写入目标） / Internal phase
    _eFaultFrom: E_DL_MpvPhase := E_DL_MpvPhase.eIdle;    // 故障来源相（锁存量） / Faulting phase, latched
    _eCause    : E_DL_MpvCause := E_DL_MpvCause.eNone;    // 成因锁存量 / Latched cause
    tonEvacTo  : TON;           // 抽真空相专用超时，段 0 无条件调用 / Evacuation dedicated timeout
    tonHoldTo  : TON;           // 真空保持相专用时长，段 0 无条件调用 / Hold dedicated duration
    tonBreakTo : TON;           // 破空相专用超时，段 0 无条件调用 / Air-break dedicated timeout
    tonReliefTo: TON;           // 泄压相专用时长，段 0 无条件调用 / Relief dedicated duration
    rtStart    : R_TRIG;        // 启动沿实例，段 0 无条件调用 / Start edge instance
    rtReset    : R_TRIG;        // 复位沿实例，段 0 无条件调用 / Reset edge instance
    rtVacIn    : R_TRIG;        // 真空到位沿实例，段 0 无条件调用 / Vacuum-reached edge instance
    rtBreakIn  : R_TRIG;        // 破空到位沿实例，段 0 无条件调用 / Break-done edge instance
    _bVacSeen  : BOOL;          // 真空到位沿锁存（进相清、捕获沿置位） / Vacuum-reached edge latch
    _bBreakSeen: BOOL;          // 破空到位沿锁存（进相清、捕获沿置位） / Break-done edge latch
    _bFault    : BOOL;          // 故障锁存位（锁存量） / Latched fault bit
    _bCfgBad   : BOOL;          // 组态非法当拍量 [-] / Illegal configuration this scan
    _bBusyPrev : BOOL;          // 上拍忙碌快照（用于完成脉冲） / Busy snapshot for the completion pulse
END_VAR

(* —— 段 0：组态闸 + 四枚专用 TON 与两枚沿无条件周期刷新 —— *)
_bCfgBad := (tEvac <= T#0S) OR (tHold <= T#0S)                  // 抽真空/保持时长须为正 / Evacuation and hold durations must be positive
         OR (tBreak <= T#0S) OR (tRelief <= T#0S);              // 破空/泄压时长须为正 / Break and relief durations must be positive
rtStart(CLK := bStart);                                          // 启动沿，每拍必调（R228A） / Start edge, every scan
rtReset(CLK := bReset);                                          // 复位沿，每拍必调 / Reset edge, every scan
rtVacIn(CLK := bVacReached);                                     // 真空到位沿，每拍必调 / Vacuum-reached edge, every scan
rtBreakIn(CLK := bBreakDone);                                    // 破空到位沿，每拍必调 / Break-done edge, every scan
tonEvacTo(IN := (_eState = E_DL_MpvPhase.eEvac), PT := tEvac);        // 抽真空相专用超时（进相计时，出相自复位） / Evacuation dedicated timeout
tonHoldTo(IN := (_eState = E_DL_MpvPhase.eHold), PT := tHold);        // 保持相专用时长 / Hold dedicated duration
tonBreakTo(IN := (_eState = E_DL_MpvPhase.eBreak), PT := tBreak);     // 破空相专用超时 / Air-break dedicated timeout
tonReliefTo(IN := (_eState = E_DL_MpvPhase.eRelief), PT := tRelief);  // 泄压相专用时长 / Relief dedicated duration

(* —— 段 1：单拍量预清零（锁存量 _eFaultFrom/_eCause/_bFault/_bBusyPrev 不入清单，R107） —— *)
bEvacActive   := FALSE;     // 抽真空相指示预清 / Evacuation indicator preset
bHoldActive   := FALSE;     // 保持相指示预清 / Hold indicator preset
bBreakActive  := FALSE;     // 破空相指示预清 / Break indicator preset
bReliefActive := FALSE;     // 泄压相指示预清 / Relief indicator preset
bBusy         := FALSE;     // 忙碌指示预清 / Busy preset
bComplete     := FALSE;     // 完成脉冲预清 / Complete pulse preset
bAborted      := FALSE;     // 中止脉冲预清 / Aborted pulse preset
bError        := FALSE;     // 故障标志预清（R45 配对） / Error flag preset

(* —— 段 2：组态闸（相时间非正即故障，记录来源相） —— *)
IF _bCfgBad THEN
    IF _eState <> E_DL_MpvPhase.eFault THEN
        _eFaultFrom := _eState;                         // 记录跌入故障时所在相 / Record the phase that faulted
    END_IF
    _bFault := TRUE;                                    // 锁存 / Latch
    _eCause := E_DL_MpvCause.eCfgIllegal;               // 归因：组态非法 / Cause: illegal configuration
    _eState := E_DL_MpvPhase.eFault;                    // 入故障相 / Enter fault phase
END_IF

(* —— 段 3：迁出链（bReset 上升沿 或 bStop 停机优先；两条都显式写出，R228B） —— *)
IF rtReset.Q THEN
    _bFault     := FALSE;                               // 清故障锁存 / Clear the fault latch
    _eCause     := E_DL_MpvCause.eNone;                 // 清成因 / Clear cause
    _eFaultFrom := E_DL_MpvPhase.eIdle;                 // 清来源相 / Clear the faulting phase
    _bVacSeen   := FALSE;                               // 清真空到位锁存（迁出链防残留，R310/R311） / Clear vacuum latch on exit chain
    _bBreakSeen := FALSE;                               // 清破空到位锁存（迁出链防残留，R310/R311） / Clear break latch on exit chain
    _eState     := E_DL_MpvPhase.eIdle;                 // 回待机相（迁出路径 1） / Back to idle, exit path 1
END_IF
IF bStop AND (_eState <> E_DL_MpvPhase.eIdle) THEN
    bAborted := TRUE;                                   // 中止脉冲 / Abort pulse
    IF _eState = E_DL_MpvPhase.eFault THEN
        _bFault := FALSE;                               // 停机优先：故障相也允许被停机清出 / Stop wins, clears even the fault
        _eCause := E_DL_MpvCause.eNone;                 // 清成因 / Clear cause
    END_IF
    _eFaultFrom := E_DL_MpvPhase.eIdle;                 // 清来源相 / Clear the faulting phase
    _bVacSeen   := FALSE;                               // 清真空到位锁存（迁出链防残留） / Clear vacuum latch on exit chain
    _bBreakSeen := FALSE;                               // 清破空到位锁存（迁出链防残留） / Clear break latch on exit chain
    _eState     := E_DL_MpvPhase.eIdle;                 // 回待机相（迁出路径 2） / Back to idle, exit path 2
END_IF

(* —— 段 4：顺控相迁移（只在无故障时推进；每相出口条件显式成对） —— *)
IF (NOT _bFault) AND (NOT _bCfgBad) AND (NOT bStop) THEN
    CASE _eState OF

    E_DL_MpvPhase.eIdle:
        IF rtStart.Q THEN
            _bVacSeen := FALSE;                                 // 进相首拍清到位锁存（防跨循环残留） / Clear vacuum latch on phase entry
            _eState := E_DL_MpvPhase.eEvac;                     // 启动沿入抽真空相 / Start edge enters evacuation
        END_IF

    E_DL_MpvPhase.eEvac:
        IF rtVacIn.Q THEN
            _bVacSeen := TRUE;                                  // 捕获真空到位沿并锁存（脉冲型兼容） / Capture vacuum-reached edge into latch
        END_IF
        IF tonEvacTo.Q AND _bVacSeen THEN
            _eState := E_DL_MpvPhase.eHold;                     // 定时到 ∧ 真空到位锁存：进保持相 / Timer done and vacuum latch set
        ELSIF tonEvacTo.Q AND (NOT _bVacSeen) THEN
            _eFaultFrom := E_DL_MpvPhase.eEvac;                 // 记录故障来源相 / Record the faulting phase
            _bFault := TRUE;                                    // 锁存 / Latch
            _eCause := E_DL_MpvCause.eVacTimeout;               // 归因：抽真空超时 / Cause: evacuation timeout
            _eState := E_DL_MpvPhase.eFault;                    // 入故障相 / Enter fault phase
        END_IF

    E_DL_MpvPhase.eHold:
        IF tonHoldTo.Q THEN
            _bBreakSeen := FALSE;                               // 进破空相首拍清到位锁存（防跨循环残留） / Clear break latch on phase entry
            _eState := E_DL_MpvPhase.eBreak;                    // 保持时长到：进破空相 / Hold done enters air break
        END_IF

    E_DL_MpvPhase.eBreak:
        IF rtBreakIn.Q THEN
            _bBreakSeen := TRUE;                                // 捕获破空到位沿并锁存（脉冲型兼容） / Capture break-done edge into latch
        END_IF
        IF tonBreakTo.Q AND _bBreakSeen THEN
            _eState := E_DL_MpvPhase.eRelief;                   // 定时到 ∧ 破空到位锁存：进泄压相 / Timer done and break latch set
        ELSIF tonBreakTo.Q AND (NOT _bBreakSeen) THEN
            _eFaultFrom := E_DL_MpvPhase.eBreak;                // 记录故障来源相 / Record the faulting phase
            _bFault := TRUE;                                    // 锁存 / Latch
            _eCause := E_DL_MpvCause.eBreakTimeout;             // 归因：破空超时 / Cause: air-break timeout
            _eState := E_DL_MpvPhase.eFault;                    // 入故障相 / Enter fault phase
        END_IF

    E_DL_MpvPhase.eRelief:
        IF tonReliefTo.Q THEN
            _eState := E_DL_MpvPhase.eIdle;                     // 泄压完成：回待机相 / Relief done returns to idle
        END_IF

    E_DL_MpvPhase.eFault:
        ;                                                       // 故障相：由段 3 两条迁出路径处理 / Handled by the two exit paths in stage 3

    ELSE
        _eFaultFrom := _eState;                                 // 记录异常相 / Record the anomalous phase
        _eCause := E_DL_MpvCause.ePhaseBad;                     // 归因：非法相位 / Cause: illegal phase
        _bFault := TRUE;                                        // 锁存 / Latch
        _eState := E_DL_MpvPhase.eFault;                        // 强拉故障相 / Force fault phase

    END_CASE
END_IF

(* —— 段 5：完成脉冲（由"忙碌→空闲"且无中止无故障的沿派生，单拍） —— *)
IF _bBusyPrev AND (_eState = E_DL_MpvPhase.eIdle) AND (NOT bAborted) AND (NOT _bFault) THEN
    bComplete := TRUE;                                          // 四相走完 / All four phases finished
END_IF
_bBusyPrev := (_eState <> E_DL_MpvPhase.eIdle) AND (_eState <> E_DL_MpvPhase.eFault);   // 忙碌快照（本拍末） / Busy snapshot at body end

(* —— 段 6：出口单点映射（相指示与相别同源，R191） —— *)
bEvacActive   := (_eState = E_DL_MpvPhase.eEvac);               // 抽真空相指示 / Evacuation indicator
bHoldActive   := (_eState = E_DL_MpvPhase.eHold);               // 保持相指示 / Hold indicator
bBreakActive  := (_eState = E_DL_MpvPhase.eBreak);              // 破空相指示 / Break indicator
bReliefActive := (_eState = E_DL_MpvPhase.eRelief);             // 泄压相指示 / Relief indicator
bBusy         := (_eState <> E_DL_MpvPhase.eIdle) AND (_eState <> E_DL_MpvPhase.eFault);   // 忙碌 / Busy
bError        := _bFault OR _bCfgBad;                           // 故障标志 = 锁存或组态非法 / Error = latch or illegal config
ePhase        := _eState;                                       // 当前相出口 / Present phase outlet
eFaultFrom    := _eFaultFrom;                                   // 故障来源相出口 / Faulting phase outlet
eCause        := _eCause;                                       // 成因出口 / Cause outlet

END_FUNCTION_BLOCK

(* ---- FB_DL_MoldCoolingZoneSeq.st ---- *)
(*==============================================================================
 * 组件名称 (Component)  : FB_DL_MoldCoolingZoneSeq
 * 所属子库 (Sublibrary) : DL_Process
 * 当前版本 (Version)    : 1.0.1
 * 兼容性   (Platform)   : CODESYS 3.5 / TwinCAT 3 / 汇川 InoProShop / 施耐德 Machine Expert
 *                         仅依赖 IEC 61131-3 标准库（TON / R_TRIG / ABS / MAX / SHL）
 * 功能描述 (Function)   : 注塑模具分区冷却时序控制：
 *                         eIdle → ePreHeat（预热到 fTempSet 的 ±fTempTol 内并驻留 tHeatDwell）
 *                         → eZoneFlow（按 iZoneCount 逐区开阀，逐区确认流量开关）→
 *                         eBalance（各区温差 ≤ fBalTol 且持续 tBalTime）→ eBlow（吹扫
 *                         tBlowTime）→ eDone；任一分区流量在 tFlowTimeout 内未确认 →
 *                         **eDegraded**（该区阀关闭并置 iFaultZoneMask 对应位，其余分区
 *                         继续依次开启，整段流程不中断）；急停 bEStop 或模温超上限
 *                         bMoldTempHigh → **eFault** 当拍全阀关（出口侧再以 bFaultCut 双保险）。
 * 接口     (Interface)  : 输入 17 项（启动/复位/急停/模温上限/模温/预热设定/容差/
 *                         预热驻留/分区数/8 路流量反馈/8 路分区温度/流量超时/平衡容差/
 *                         平衡持续/吹扫时长），输出 7 项（状态回执/8 路阀/吹扫阀/故障分区
 *                         位图/完成/降级/故障与码）。
 * 边界     (Boundary)   : ① 分区数 iZoneCount 钳位到 1..8；数组下标在每次访问前用
 *                            整数域闸保护（R4 下标钳位），越界即不访问。
 *                         ② 流量超时只降级不中止：置位图、关该区阀、继续其余分区；
 *                            全部区均超时仍走 eBalance → eBlow → eDone（流程闭环）。
 *                         ③ 急停与模温上限为最高优先级拦截，位于 CASE 之前；出口侧
 *                            bFaultCut 再做一次硬件切断（双保险）。
 *                         ④ fMoldTemp / 分区温度非有限值按「判据不可满足」处理
 *                            （不假装通过），并在温度类判据中显式披露。
 *                         ⑤ 零全局耦合（无 GVL / VAR_EXTERNAL / %I / %Q）。
 * 码表     (Codes)      : 本件占用 16#0004_1010 ~ 16#0004_101F 区间，实际使用 7 个：
 *                         1010 信息级 分区数越界已钳位；1011 信息级 某分区流量超时已降级；
 *                         1012 故障级 急停动作；1013 故障级 模温超上限；
 *                         1014 故障级 模温反馈非有限；1015 故障级 非法状态兜底；
 *                         1016 信息级 平衡温差长期不收敛，按超时降级进吹扫。
 *                         信息级码永不置 bError；故障级码锁存回放，bReset 且条件消失解除。
 * 分工声明 (Scope)      : 本件只做「分区冷却时序 + 阀位排列」，不做温度 PID 调节
 *                         （温度闭环归 FB_DL_TempPidZone 类组件），不做流量计标定。
 * 开源溯源 (Origin)     : 开源溯源：原创实现（无外部代码引入）
 * 红线自检 (Redline)    : R1 ✓ 零 GVL / VAR_EXTERNAL ｜ R2 ✓ 零 %I/%Q/%M
 *                         R3 ✓ 纯 IEC 61131-3 ｜ R4 ✓ 下标钳位 + 非有限双判 + 容差 1E-9
 *                         R5 ✓ 声明逐行同行双语注释 ｜ R6 ✓ 八态 ENUM + CASE + ELSE
 *                         R7 ✓ 五个定时器/边沿实例全部无条件每周期调用
 * 修订历史 (Revision)   : 2026-11-23  v1.0.0  R77 首版
 *                         2026-11-23  v1.0.1  R77 闸修复（Inf 阈值直比 / eFault 复位出口 / eBalance 超时兜底）
 * 验收向量 (Acceptance) :
 *   V1 bStart 上升、模温 25 ℃、fTempSet=80 ℃：eStateOut=ePreHeat，8 路阀全 FALSE；
 *      模温升至 80 ℃（容差 2 ℃）后驻留 tHeatDwell，随后 eStateOut=eZoneFlow。
 *   V2 iZoneCount=3、三区流量开关在 1s 内依次闭合：eStateOut 依次 eZoneFlow(区1→2→3)
 *      → eBalance → eBlow → eDone，iFaultZoneMask=0，bDone=TRUE。
 *   V3 iZoneCount=3、区 2 流量开关始终不闭合（tFlowTimeout=10s）：
 *      10s 后 iFaultZoneMask 第 2 位 = 1（十进制 2）、abZoneValve[2]=FALSE、
 *      eStateOut=eDegraded，区 3 仍被开启；后续进入 eBalance → eBlow → eDone，bDegraded=TRUE。
 *   V4 任何状态 bEStop 上升：当拍 eStateOut=eFault、8 路阀与吹扫阀全 FALSE、
 *      uErrorId=16#0004_1012、bError=TRUE；bReset 且 bEStop 回落才回 eIdle。
 *   V5 任何状态 bMoldTempHigh 上升：当拍 eStateOut=eFault、全阀关、
 *      uErrorId=16#0004_1013；fMoldTemp=NaN 时 uErrorId=16#0004_1014 且不进入 ePreHeat。
 *   V6（R77 闸补）bEStop 触发进 eFault 后保持 bEStop=FALSE、bReset 保持一拍 →
 *      eStateOut 回归 eIdle，bFaultCut 落 FALSE，bError=FALSE（eFault 唯一出口可到达）。
 *   V7（R77 闸补）eBalance 内分区温差长期大于 fBalTol（tonBal 永不 Q）→ 超过
 *      tBalTime×5 后 eStateOut=eBlow、uErrorId=16#0004_1016、bError=FALSE（信息级降级）。
 *============================================================================*)

(*-----------------------------------------------------------------------------
 * 调用示例 (Instance guide)：
 *   声明于调用方 FB 的 VAR 区：fbCool : FB_DL_MoldCoolingZoneSeq;
 *   每周期无条件调用：fbCool(bStart := xMoldStart, bReset := xReset,
 *                            bEStop := xEStopSafe, bMoldTempHigh := xTempHiAlarm,
 *                            fMoldTemp := stMold.fTemp, fTempSet := rTempSp,
 *                            iZoneCount := nZoneNum);
 *   数组引脚：abFlowFb / afZoneTemp 直接指向上层结构体中的 8 元数组。
 *   出口用法：abZoneValve 逐路驱动电磁阀，bFaultCut 由本件内部消费，无需使用者再 AND。
 *   调参指引：tFlowTimeout 取流量开关响应时间的 3 倍；fBalTol 取工艺允许温差的一半；
 *            tBlowTime 取管路容积 ÷ 吹扫流量再加 2 s 余量。
 *----------------------------------------------------------------------------*)

(*-----------------------------------------------------------------------------
 * 枚举: E_DL_MczState（归属 DL_Process，与 FB_DL_MoldCoolingZoneSeq 同文件）
 * 含义: 模具分区冷却时序状态机的离散状态。正序为 eIdle → ePreHeat → eZoneFlow →
 *       eBalance → eBlow → eDone；eDegraded 为「降级继续」分支相，eFault 为安全相。
 *----------------------------------------------------------------------------*)
TYPE E_DL_MczState :
(
    eIdle     := 0,    // 空闲态：全阀关，等 bStart 上升沿 / Idle: all valves closed, waiting for bStart rise
    ePreHeat  := 10,   // 预热态：等模温进入 设定±容差 并驻留 tHeatDwell / Pre-heat: wait for mould temperature in band plus dwell
    eZoneFlow := 20,   // 分区开阀态：按 iZone 逐区开阀并确认流量反馈 / Zone flow: open valve by index and confirm flow feedback
    eBalance  := 30,   // 平衡态：各区温差 ≤ fBalTol 持续 tBalTime / Balance: zone temperature spread within tolerance for tBalTime
    eBlow     := 40,   // 吹扫态：全分区阀关、吹扫阀开 tBlowTime / Blow: zone valves closed, blow valve open for tBlowTime
    eDone     := 50,   // 完成态：全阀关，保持完成标志直到 bStart 跌落 / Done: all valves closed, holds until bStart falls
    eDegraded := 60,   // 降级态：某区流量超时，该区已关阀置位图，其余分区继续 / Degraded: one zone failed, others keep sequencing
    eFault    := 99    // 故障安全态：急停/模温超上限/非法状态，全阀立即关 / Fault safe state: e-stop or over-temperature, all valves closed at once
);
END_TYPE

(*==============================================================================
 * 功能块: FB_DL_MoldCoolingZoneSeq
 * 调用约定: 每周期无条件调用一次；五个定时器/边沿实例在段 2 无条件刷新。
 * 出口语义: abZoneValve / bBlowValve 在 eFault（或急停、模温超上限）当拍即被强制关断，
 *           不依赖状态机内部清零是否已执行（双保险）。
 *============================================================================*)
FUNCTION_BLOCK FB_DL_MoldCoolingZoneSeq
VAR_INPUT
    bStart        : BOOL := FALSE;      // 启动（上升沿开始流程，跌落回 eIdle）/ Start, rising edge begins the sequence, falling returns to eIdle
    bReset        : BOOL := FALSE;      // 复位（电平有效），解除故障锁存 / Reset (level), clears the fault latch
    bEStop        : BOOL := FALSE;      // 急停信号，TRUE = 急停动作，最高优先级拦截 / Emergency stop, TRUE = actuated, highest priority interlock
    bMoldTempHigh : BOOL := FALSE;      // 模温超上限开关，TRUE = 超限，最高优先级拦截 / Mould over-temperature switch, TRUE = over limit, highest priority
    fMoldTemp     : REAL := 0.0;        // 模具当前温度 [℃] / Current mould temperature [degC]
    fTempSet      : REAL := 80.0;       // 预热设定温度 [℃] / Pre-heat setpoint temperature [degC]
    fTempTol      : REAL := 2.0;        // 预热到温容差 [℃] / Pre-heat in-band tolerance [degC]
    tHeatDwell    : TIME := T#10S;      // 到温驻留时间 [s] / Dwell time after reaching temperature [s]
    iZoneCount    : INT := 4;           // 参与时序的分区数，钳位 1..8 [-] / Number of zones in the sequence, clamped 1..8
    abFlowFb      : ARRAY[1..8] OF BOOL;      // 分区流量开关反馈，TRUE = 有流量 [BOOL] / Per-zone flow switch feedback, TRUE = flow present
    afZoneTemp    : ARRAY[1..8] OF REAL;      // 分区冷却水温反馈 [℃] / Per-zone coolant temperature feedback [degC]
    tFlowTimeout  : TIME := T#10S;      // 单区流量确认超时 [s] / Per-zone flow confirmation timeout [s]
    fBalTol       : REAL := 3.0;        // 平衡温差容差 [℃] / Balance temperature spread tolerance [degC]
    tBalTime      : TIME := T#15S;      // 平衡持续确认时间 [s] / Balance confirmation duration [s]
    tBlowTime     : TIME := T#5S;       // 吹扫时长 [s] / Blow duration [s]
END_VAR
VAR_OUTPUT
    eStateOut     : E_DL_MczState;      // 状态机当前状态回执 [-] / Current state feedback
    abZoneValve   : ARRAY[1..8] OF BOOL;      // 分区冷却阀输出，TRUE = 开阀 [BOOL] / Per-zone coolant valve output, TRUE = open
    bBlowValve    : BOOL;               // 吹扫阀输出，TRUE = 开 / Blow valve output, TRUE = open
    iFaultZoneMask: INT;                // 流量超时分区位图，位 0 = 1 区 [-] / Zone fault bitmap, bit 0 = zone 1
    bDone         : BOOL;               // 流程完成标志（eDone 相保持）/ Sequence done flag, held during eDone
    bDegraded     : BOOL;               // 降级运行标志（至少一区流量超时）/ Degraded run flag, at least one zone timed out
    bFaultCut     : BOOL;               // 强制切断回执，TRUE 表示出口已被安全侧切断 / Forced cut-off feedback, TRUE means outlets are cut by the safety side
    bValid        : BOOL;               // 出口数据可信标志 / Output data trustworthy flag
    bError        : BOOL;               // 故障级标志，与 uErrorId 严格联动 / Fault-level flag, strictly coupled with uErrorId
    uErrorId      : UDINT;              // 错误码，0 = 无码 / Error code, 0 = no code
END_VAR
VAR
    eState        : E_DL_MczState;      // 内部状态 [-] / Internal state
    tonHeat       : TON;                // 到温驻留定时器，无条件刷新 / In-band dwell timer, refreshed unconditionally
    tonFlow       : TON;                // 单区流量确认定时器，无条件刷新 / Per-zone flow confirmation timer, refreshed unconditionally
    tonBal        : TON;                // 平衡持续定时器，无条件刷新 / Balance duration timer, refreshed unconditionally
    tonBlow       : TON;                // 吹扫时长定时器，无条件刷新 / Blow duration timer, refreshed unconditionally
    tonBalTmo     : TON;                // 平衡超时兜底定时器（tBalTime×5），无条件刷新 / Balance timeout watchdog timer, refreshed unconditionally
    rtrStart      : R_TRIG;             // 启动上升沿检测，无条件刷新 / Start rising edge detector, refreshed unconditionally
    abZoneOn      : ARRAY[1..8] OF BOOL;      // 分区阀内部指令锁存 [BOOL] / Internal per-zone valve command latch
    iZone         : INT;                // 当前处理分区号，1 基 [-] / Current zone index, one based
    iZonePrev     : INT;                // 上一拍分区号，用于换区复位定时器 [-] / Previous zone index, used to restart the flow timer
    iZoneUse      : INT;                // 钳位后的实际分区数 [-] / Clamped effective zone count
    iIdx          : INT;                // 通用循环下标 [-] / Generic loop index
    bZoneNew      : BOOL;               // 换区单拍标志（新分区首拍）/ Zone-changed single-shot flag, first scan of a new zone
    bFlowOk       : BOOL;               // 当前分区流量已确认 / Current zone flow confirmed
    bTempInBand   : BOOL;               // 模温已进入设定带 [-]/[℃] / Mould temperature inside the band
    bTempFinite   : BOOL;               // 模温反馈为有限值 / Mould temperature feedback is finite
    bZoneTempOk   : BOOL;               // 全部分区温度均有限且可比 / All active zone temperatures finite and comparable
    bSpreadOk     : BOOL;               // 分区温差在容差内 / Zone temperature spread inside tolerance
    bFaultLatch   : BOOL;               // 安全故障锁存位 / Safety fault latch
    bFaultCond    : BOOL;               // 安全故障条件（急停或模温超上限）/ Safety fault condition, e-stop or over-temperature
    bCountClamped : BOOL;               // 分区数被钳位的单拍记录 / Zone count clamp record
    wBitTmp       : WORD;               // 位图构造中间量 [位图] / Bitmap construction scratch [bitmap]
    nShift        : INT;                // 移位量，恒 ≤ 7，绝不等于位宽 [位] / Shift amount, always <= 7, never equals bit width [bit]
    fZoneMax      : REAL;               // 活动分区最高水温 [℃] / Highest coolant temperature among active zones [degC]
    fZoneMin      : REAL;               // 活动分区最低水温 [℃] / Lowest coolant temperature among active zones [degC]
    fTempTolEff   : REAL;               // 钳位后到温容差 [℃] / Clamped in-band tolerance [degC]
    fBalTolEff    : REAL;               // 钳位后平衡容差 [℃] / Clamped balance tolerance [degC]
    uInfoCode     : UDINT;              // 信息级码暂存 / Info-level code scratch
END_VAR
VAR CONSTANT
    DL_MCZ_ZONE_MAX : INT := 8;                    // 分区数硬上限（数组上界）[-] / Hard zone limit, the array upper bound
    DL_MCZ_ZONE_MIN : INT := 1;                    // 分区数硬下限 [-] / Hard zone lower bound
    DL_MCZ_BIT_ONE  : WORD := 16#0001;             // 位图起始掩码（1 区）/ Bitmap base mask for zone one
    DL_MCZ_WORD_0   : WORD := 16#0000;             // 零哨兵，避免裸字面量比较 / Zero sentinel avoiding bare literal comparison
    DL_MCZ_TOL      : REAL := 1.0E-3;              // 容差下限硬钳位值 [℃] / Tolerance lower clamp value [degC]
    DL_MCZ_EPS      : REAL := 1.0E-9;              // 浮点比较容差（统一口径）/ Unified floating point comparison tolerance
    DL_MCZ_ZERO     : REAL := 0.0;                 // 零基准哨兵 / Zero reference sentinel
    DL_MCZ_OK       : UDINT := 16#0000_0000;       // 无码哨兵 / No-code sentinel
    DL_MCZ_RMAX     : REAL := 3.4028235E38;         // 本机 REAL 可表示上限，Inf 阈值直比基准 [无量纲] / Locally representable REAL maximum, Inf threshold base
    DL_MCZ_BAL_TMO_FACTOR : INT := 5;               // 平衡超时倍率，超时 = tBalTime × 本倍率 [-] / Balance timeout factor, timeout = tBalTime x this
END_VAR

(*------------------------------------------------------------------------------
 * 段 0｜参数域闸（不中断扫描）：分区数钳位 1..8、容差下限钳位
 *      Parameter domain gate: clamp zone count to 1..8 and tolerance floors
 *-----------------------------------------------------------------------------*)
uInfoCode  := DL_MCZ_OK;                                    // 信息码预置无码 / Preset no info code
bCountClamped := FALSE;                                     // 钳位记录预置 / Preset clamp record FALSE

IF iZoneCount < DL_MCZ_ZONE_MIN THEN
    iZoneUse      := DL_MCZ_ZONE_MIN;                       // 分区数过小钳到 1 / Too few zones clamped to one
    bCountClamped := TRUE;                                  // 记录钳位 / Record the clamp
ELSIF iZoneCount > DL_MCZ_ZONE_MAX THEN
    iZoneUse      := DL_MCZ_ZONE_MAX;                       // 分区数过大钳到 8（数组上界）/ Too many zones clamped to eight
    bCountClamped := TRUE;                                  // 记录钳位 / Record the clamp
ELSE
    iZoneUse := iZoneCount;                                 // 合法分区数原值生效 / Legal zone count applied as-is
END_IF
IF bCountClamped THEN
    uInfoCode := 16#0004_1010;                              // 信息级：分区数越界已钳位 / Info: zone count out of range, clamped
END_IF

fTempTolEff := MAX(fTempTol, DL_MCZ_TOL);                   // 到温容差下限钳位 [℃] / In-band tolerance floor [degC]
fBalTolEff  := MAX(fBalTol, DL_MCZ_TOL);                    // 平衡容差下限钳位 [℃] / Balance tolerance floor [degC]

(*------------------------------------------------------------------------------
 * 段 1｜判据量计算：模温带判定（非有限值判「不可满足」）与当前分区流量确认
 *      Predicate computation: temperature band test treating non-finite as unsatisfied
 *-----------------------------------------------------------------------------*)
bTempFinite := NOT ((fMoldTemp <> fMoldTemp)
                    OR (fMoldTemp > DL_MCZ_RMAX) OR (fMoldTemp < -DL_MCZ_RMAX));          // 模温有限判定：NaN 自反 + Inf 阈值直比 / Finite test: NaN self-comparison plus Inf threshold
bTempInBand := bTempFinite AND (ABS(fMoldTemp - fTempSet) <= fTempTolEff);                 // 到温带判定 [℃] / In-band test [degC]

bFlowOk := FALSE;                                           // 默认未确认流量 / Flow not confirmed by default
IF (iZone >= DL_MCZ_ZONE_MIN) AND (iZone <= DL_MCZ_ZONE_MAX) THEN
    bFlowOk := abFlowFb[iZone];                             // 下标域闸通过才访问数组 / Array accessed only after the index gate
END_IF

bZoneNew := iZone <> iZonePrev;                             // 换区单拍标志（本拍为新分区首拍）/ Zone change single shot

(*------------------------------------------------------------------------------
 * 段 2｜定时器与边沿实例无条件刷新（红线 R7）：全部置于 CASE 之外
 *      Unconditional refresh of timers and edge detectors, all outside the CASE
 *      流量窗口 IN 串 NOT bZoneNew：换区当拍强制复位 ET，绝不让上一区余量带入新区
 *-----------------------------------------------------------------------------*)
rtrStart(CLK := bStart);                                    // 启动上升沿，无条件调用 / Start edge, called unconditionally

tonHeat(IN := bTempInBand AND (eState = ePreHeat), PT := tHeatDwell);   // 到温驻留计时，无条件调用 / In-band dwell timer, called unconditionally

tonFlow(IN := ((eState = eZoneFlow) OR (eState = eDegraded))
             AND (iZone >= DL_MCZ_ZONE_MIN) AND (iZone <= iZoneUse)
             AND (NOT bFlowOk) AND (NOT bZoneNew), PT := tFlowTimeout);   // 单区流量窗，无条件调用 / Zone flow window, called unconditionally

tonBal(IN := bSpreadOk AND (eState = eBalance), PT := tBalTime);        // 平衡持续计时，无条件调用 / Balance duration timer, called unconditionally

tonBlow(IN := (eState = eBlow), PT := tBlowTime);                       // 吹扫时长计时，无条件调用 / Blow duration timer, called unconditionally

tonBalTmo(IN := (eState = eBalance), PT := tBalTime * DL_MCZ_BAL_TMO_FACTOR);   // 平衡超时兜底计时，IN 挂状态量故离相即自复位，无条件调用 / Balance watchdog, self-reset by leaving the state, called unconditionally

(*------------------------------------------------------------------------------
 * 段 3｜安全拦截（最高优先级，位于 CASE 之前）：急停 / 模温超上限 → 当拍进 eFault
 *      Safety interlock before the CASE: e-stop or over-temperature enters eFault at once
 *      故障锁存解除路径唯一：bReset 且 bEStop 回落 且 bMoldTempHigh 回落
 *      解除当拍状态同步回归 eIdle（eFault 的唯一出口，须在段 4 之前生效，否则永久停故障态）
 *      Sole clear path: reset with both conditions gone; the same scan returns the state
 *      machine to eIdle, which is the only exit from eFault, applied before segment 4.
 *-----------------------------------------------------------------------------*)
bFaultCond := bEStop OR bMoldTempHigh;                      // 安全故障条件 / Safety fault condition

IF bFaultCond THEN
    bFaultLatch := TRUE;                                    // 安全故障锁存置位 / Safety fault latch set
    eState      := eFault;                                   // 当拍强制进安全相 / Force the safe state this scan
ELSIF bFaultLatch THEN
    IF bReset THEN
        bFaultLatch := FALSE;                               // 唯一解除路径：复位且条件已回落 / Sole clear path: reset with conditions gone
        eState      := eIdle;                               // 复位回归怠速态：eFault 的唯一出口（段 4 之前生效）/ Reset returns to idle, the only exit from eFault, applied before segment 4
    ELSE
        eState := eFault;                                   // 未复位则保持安全相 / Stay in the safe state without reset
    END_IF
END_IF

(*------------------------------------------------------------------------------
 * 段 4｜主状态机（红线 R6）：ENUM + CASE + ELSE 兜底
 *      Main state machine with enum, case coverage and ELSE interception
 *      迁入安全相后的出口清零由段 5 的 bFaultCut 统一保证，CASE 内不重复做门控
 *-----------------------------------------------------------------------------*)
IF eState = eFault THEN
    (* 安全相出口：分区阀指令全部清零（CASE 内不做二次判定，避免同拍竞态）*)
    (* Safe state outlets: clear every zone command, no second judgement to avoid race *)
    FOR iIdx := DL_MCZ_ZONE_MIN TO DL_MCZ_ZONE_MAX DO
        abZoneOn[iIdx] := FALSE;                            // 逐路清指令 / Clear command zone by zone
    END_FOR
    iZone  := DL_MCZ_ZONE_MIN;                              // 分区游标回 1 / Zone cursor back to one
    bDone  := FALSE;                                        // 完成标志清除 / Done flag cleared
    bValid := FALSE;                                        // 出口数据不可信 / Outlet data untrustworthy
ELSE
    CASE eState OF

        eIdle:
            (* 空闲：游标与位图复位，等 bStart 上升沿 *)
            (* Idle: reset cursor and bitmap, wait for the start edge *)
            FOR iIdx := DL_MCZ_ZONE_MIN TO DL_MCZ_ZONE_MAX DO
                abZoneOn[iIdx] := FALSE;                    // 逐路清阀指令 / Clear valve command zone by zone
            END_FOR
            iZone          := DL_MCZ_ZONE_MIN;              // 游标回 1 / Cursor back to one
            iFaultZoneMask := 0;                            // 位图清零 / Bitmap cleared
            bDone          := FALSE;                        // 完成标志清除 / Done flag cleared
            bDegraded      := FALSE;                        // 降级标志清除 / Degraded flag cleared
            bValid         := TRUE;                         // 空闲相出口可信 / Outlets trustworthy in idle
            IF rtrStart.Q AND (NOT bTempFinite) THEN
                eState := eFault;                           // 温度反馈已坏：拒绝启动（不漏判）/ Broken feedback, refuse to start
            ELSIF rtrStart.Q THEN
                eState := ePreHeat;                         // 启动沿进预热 / Start edge enters pre-heat
            END_IF

        ePreHeat:
            (* 预热：到温带内驻留 tHeatDwell 后进入分区开阀；进相前温度坏值转故障 *)
            (* Pre-heat: dwell in band, then go to zone flow, broken feedback turns to fault *)
            FOR iIdx := DL_MCZ_ZONE_MIN TO DL_MCZ_ZONE_MAX DO
                abZoneOn[iIdx] := FALSE;                    // 预热相不开分区阀 / No zone valve open during pre-heat
            END_FOR
            bValid := TRUE;                                 // 预热相出口可信 / Outlets trustworthy in pre-heat
            IF NOT bTempFinite THEN
                eState := eFault;                           // 温度非有限：进安全相 / Non-finite temperature, safe state
            ELSIF NOT bStart THEN
                eState := eIdle;                            // 启动撤销回空闲 / Start removed returns to idle
            ELSIF tonHeat.Q THEN
                iZone  := DL_MCZ_ZONE_MIN;                  // 到温驻留完成，游标从 1 区起 / Dwell done, cursor starts at zone one
                eState := eZoneFlow;                        // 进入分区开阀 / Enter zone flow
            END_IF

        eZoneFlow:
            (* 分区开阀：下标域闸通过才访问数组；确认 → 推进；超时 → 降级态 *)
            (* Zone flow: index gate before array access, confirm advances, timeout degrades *)
            IF iZone > iZoneUse THEN
                eState := eBalance;                         // 全部分区处理完进平衡 / All zones done, enter balance
            ELSIF iZone < DL_MCZ_ZONE_MIN THEN
                iZone := DL_MCZ_ZONE_MIN;                   // 游标防御性归位 / Defensive cursor reset
            ELSE
                abZoneOn[iZone] := TRUE;                    // 开当前分区阀 / Open the current zone valve
                bValid := TRUE;                             // 出口可信 / Outlets trustworthy
                IF bFlowOk THEN
                    iZone := iZone + 1;                     // 流量确认，推进下一区 / Flow confirmed, advance
                ELSIF tonFlow.Q THEN
                    abZoneOn[iZone] := FALSE;               // 超时先关该区阀 / Close the timed-out zone valve
                    nShift   := iZone - 1;                  // 移位量恒 0..7，绝不等于位宽 / Shift always 0..7, never the bit width
                    wBitTmp  := SHL(DL_MCZ_BIT_ONE, nShift);   // 构造该区位掩码 / Build the zone bit mask
                    IF wBitTmp <> DL_MCZ_WORD_0 THEN
                        iFaultZoneMask := iFaultZoneMask OR WORD_TO_INT(wBitTmp);   // 置位图 / Set the bitmap bit
                    END_IF
                    bDegraded := TRUE;                      // 降级标志置位 / Degraded flag set
                    uInfoCode := 16#0004_1011;              // 信息级：某区流量超时 / Info: a zone timed out
                    iZone     := iZone + 1;                 // 推进，其余分区继续 / Advance, other zones continue
                    eState    := eDegraded;                 // 进入降级相 / Enter degraded state
                END_IF
            END_IF

        eDegraded:
            (* 降级继续：与 eZoneFlow 同构但不再回头进位；超时只加位图不换相 *)
            (* Degraded continue: same body as eZoneFlow but timeouts only add bitmap bits *)
            IF iZone > iZoneUse THEN
                eState := eBalance;                         // 剩余分区处理完进平衡 / Remaining zones done, enter balance
            ELSIF iZone < DL_MCZ_ZONE_MIN THEN
                iZone := DL_MCZ_ZONE_MIN;                   // 游标防御性归位 / Defensive cursor reset
            ELSE
                abZoneOn[iZone] := TRUE;                    // 开当前分区阀 / Open the current zone valve
                bValid := TRUE;                             // 出口可信 / Outlets trustworthy
                IF bFlowOk THEN
                    iZone := iZone + 1;                     // 流量确认，推进 / Flow confirmed, advance
                ELSIF tonFlow.Q THEN
                    abZoneOn[iZone] := FALSE;               // 超时关该区阀 / Close the timed-out valve
                    nShift   := iZone - 1;                  // 移位量恒 0..7 / Shift always 0..7
                    wBitTmp  := SHL(DL_MCZ_BIT_ONE, nShift);   // 区位掩码 / Zone bit mask
                    IF wBitTmp <> DL_MCZ_WORD_0 THEN
                        iFaultZoneMask := iFaultZoneMask OR WORD_TO_INT(wBitTmp);   // 追加位图 / Add the bitmap bit
                    END_IF
                    uInfoCode := 16#0004_1011;              // 信息级：又一分区流量超时 / Info: another zone timed out
                    iZone     := iZone + 1;                 // 推进 / Advance
                END_IF
            END_IF

        eBalance:
            (* 平衡：活动分区水温极差 ≤ 容差并持续 tBalTime；阀保持开（不重写指令）*)
            (* Balance: active zone spread within tolerance for tBalTime, valves stay open *)
            bValid := TRUE;                                 // 平衡相出口可信 / Outlets trustworthy
            fZoneMax := afZoneTemp[DL_MCZ_ZONE_MIN];        // 极值初值取 1 区（下标常量，恒合法）/ Extremes start from zone one
            fZoneMin := afZoneTemp[DL_MCZ_ZONE_MIN];        // 极值初值取 1 区 / Extremes start from zone one
            bZoneTempOk := NOT ((afZoneTemp[DL_MCZ_ZONE_MIN] <> afZoneTemp[DL_MCZ_ZONE_MIN])
                             OR (afZoneTemp[DL_MCZ_ZONE_MIN] > DL_MCZ_RMAX)
                             OR (afZoneTemp[DL_MCZ_ZONE_MIN] < -DL_MCZ_RMAX));   // 首区有限判定：NaN 自反 + Inf 阈值直比 / Zone-one finite test: NaN plus Inf threshold
            FOR iIdx := DL_MCZ_ZONE_MIN TO iZoneUse DO
                IF (afZoneTemp[iIdx] <> afZoneTemp[iIdx])
                   OR (afZoneTemp[iIdx] > DL_MCZ_RMAX)
                   OR (afZoneTemp[iIdx] < -DL_MCZ_RMAX) THEN
                    bZoneTempOk := FALSE;                   // 任一区非有限即整体判据不可满足 / Any non-finite zone makes the predicate unsatisfiable
                ELSE
                    IF afZoneTemp[iIdx] > fZoneMax THEN
                        fZoneMax := afZoneTemp[iIdx];       // 更新最高水温 / Update the maximum
                    END_IF
                    IF afZoneTemp[iIdx] < fZoneMin THEN
                        fZoneMin := afZoneTemp[iIdx];       // 更新最低水温 / Update the minimum
                    END_IF
                END_IF
            END_FOR
            bSpreadOk := bZoneTempOk AND ((fZoneMax - fZoneMin) <= fBalTolEff);   // 极差判据 [℃]，非有限即不可满足 / Spread predicate [degC], unsatisfiable when non-finite
            IF NOT bStart THEN
                eState := eIdle;                            // 启动撤销回空闲 / Start removed returns to idle
            ELSIF tonBal.Q THEN
                eState := eBlow;                            // 平衡持续到，进吹扫 / Balance sustained, enter blow
            ELSIF tonBalTmo.Q THEN
                (* 温差长期不收敛按超时降级处理（信息级，不置 bError）：避免 bSpreadOk 永不成立时长期驻留且分区阀全开 *)
                (* Spread never converging degrades by timeout at info level, no bError, preventing a permanent all-valve-open dwell *)
                uInfoCode := 16#0004_1016;                  // 信息级：平衡温差长期不收敛 / Info: balance spread did not converge in time
                eState    := eBlow;                         // 保流程闭环，进吹扫 / Keep the sequence closed, enter blow
            END_IF

        eBlow:
            (* 吹扫：分区阀全关、吹扫阀开（吹扫阀由段 5 依状态派生）*)
            (* Blow: all zone valves closed, blow valve derived from the state in segment 5 *)
            FOR iIdx := DL_MCZ_ZONE_MIN TO DL_MCZ_ZONE_MAX DO
                abZoneOn[iIdx] := FALSE;                    // 吹扫前关闭全部分区阀 / Close all zone valves before blow
            END_FOR
            bValid := TRUE;                                 // 吹扫相出口可信 / Outlets trustworthy
            IF NOT bStart THEN
                eState := eIdle;                            // 启动撤销回空闲 / Start removed returns to idle
            ELSIF tonBlow.Q THEN
                eState := eDone;                            // 吹扫完成 / Blow finished
            END_IF

        eDone:
            (* 完成：全阀关，bDone 保持到 bStart 跌落 *)
            (* Done: all valves closed, bDone held until bStart falls *)
            FOR iIdx := DL_MCZ_ZONE_MIN TO DL_MCZ_ZONE_MAX DO
                abZoneOn[iIdx] := FALSE;                    // 完成相关闭全部阀 / Close all valves in the done state
            END_FOR
            bDone  := TRUE;                                 // 完成标志置位 / Done flag set
            bValid := TRUE;                                 // 完成相出口可信 / Outlets trustworthy
            IF NOT bStart THEN
                eState := eIdle;                            // 启动跌落回空闲（下一循环可重入）/ Start falls, ready for the next cycle
            END_IF

        ELSE
            (* 非法状态拦截：任何未定义枚举值一律进安全相并置兜底码 *)
            (* Illegal state interception: undefined enum values go to the safe state with a code *)
            eState    := eFault;                            // 强制回安全相 / Force the safe state
            bFaultLatch := TRUE;                            // 锁存，禁自动恢复 / Latch, no automatic recovery
            uInfoCode := 16#0004_1015;                      // 故障级：非法状态兜底 / Fault: illegal state fallback
            bValid    := FALSE;                             // 出口不可信 / Outlets untrustworthy

    END_CASE
END_IF

(*------------------------------------------------------------------------------
 * 段 5｜出口派生与安全切断（双保险）：bFaultCut = 安全相 或 急停 或 模温超上限
 *      Outlet derivation with a second safety cut, independent of state machine bookkeeping
 *-----------------------------------------------------------------------------*)
bFaultCut := bFaultCond OR (eState = eFault);               // 安全切断条件 / Safety cut-off condition
IF bFaultCut THEN
    FOR iIdx := DL_MCZ_ZONE_MIN TO DL_MCZ_ZONE_MAX DO
        abZoneOn[iIdx] := FALSE;                            // 切断时同步清指令锁存 / Clear the command latch on cut-off
    END_FOR
END_IF

FOR iIdx := DL_MCZ_ZONE_MIN TO DL_MCZ_ZONE_MAX DO
    abZoneValve[iIdx] := abZoneOn[iIdx] AND (NOT bFaultCut);   // 逐路出口映射，安全侧再 AND 一次 / Per-zone outlet mapping with a second safety AND
END_FOR
bBlowValve := (eState = eBlow) AND (NOT bFaultCut);         // 吹扫阀出口映射 / Blow valve outlet mapping

(*------------------------------------------------------------------------------
 * 段 6｜故障码统一出口（故障级锁存回放，信息级不置 bError；急停优先于超温）
 *      Unified code outlet: fault codes replayed latched, info codes never raise bError
 *-----------------------------------------------------------------------------*)
IF bFaultCond THEN
    IF bEStop THEN
        uErrorId := 16#0004_1012;                           // 故障级：急停动作 / Fault: emergency stop actuated
    ELSIF bMoldTempHigh THEN
        uErrorId := 16#0004_1013;                           // 故障级：模温超上限 / Fault: mould over-temperature
    ELSE
        uErrorId := 16#0004_1015;                           // 故障级：非法兜底 / Fault: fallback
    END_IF
    bError   := TRUE;                                       // 故障级码配对置位 / Paired fault flag set
    bValid   := FALSE;                                      // 安全相出口不可信 / Outlets untrustworthy in the safe state
ELSIF (NOT bTempFinite) AND (eState <> eIdle) THEN
    uErrorId := 16#0004_1014;                               // 故障级：模温反馈非有限 / Fault: mould temperature feedback non-finite
    bError   := TRUE;                                       // 故障级码配对置位 / Paired fault flag set
    bValid   := FALSE;                                      // 指标不可信 / Metric untrustworthy
ELSE
    uErrorId := uInfoCode;                                  // 信息级码（流量超时/分区钳位）或 0 / Info code or zero
    bError   := FALSE;                                      // 信息级不置故障标志 / Info level never raises the fault flag
END_IF

eStateOut := eState;                                        // 状态回执单一出口 / State feedback through a single outlet
iZonePrev := iZone;                                         // 换区基准刷新（本拍结束）/ Refresh the zone baseline at scan end
END_FUNCTION_BLOCK
